(* IEC 61131-3 sources: daoli-st-library/DL_Base (part 10) *)

(* ---- FB_DL_CtudEx.st ---- *)
(*==============================================================================
 * 组件名称 (Component)  : FB_DL_CtudEx
 * 所属子库 (Sublibrary) : DL_Base
 * 当前版本 (Version)    : 1.0.0
 * 兼容性   (Platform)   : CODESYS 3.5 / TwinCAT 3 / 汇川 InoProShop / Machine Expert
 *                         仅依赖 Standard.library（R_TRIG），计数本体为库内显式
 *                         判界加减法（重实现最小化：一圈判界 + 加减 1）
 * 功能描述 (Function)   : 双向计数器（CTUD）防御包装。内部以两个 R_TRIG 标准实例
 *                         分别取 bCU / bCD 上升沿，CU/CD 同拍出现时按「净额抵消法」
 *                         取净值一次性施加（net = CU沿 − CD沿，同拍加减相消不误
 *                         动作）；优先级链 bRESET > bLOAD > 计数；PV 负值钳 0；
 *                         双向饱和不回绕（达 DINT 上/下限锁定并置故障码）。
 * 溯源     (Origin)     : IEC 61131-3 标准语义的道莅防御性实现
 *                         （接口语义由 IEC 61131-3 定义，clean-room 重写，
 *                         参考公开标准条款）
 * 码位     (Diag Codes) : 信息级 16#0001_0155（本件独占）：
 *                         nPV 为负值已钳 0 ／ CU/CD 同拍抵消（净变化 0）
 *                         故障级 16#0001_0226（本件独占）：
 *                         CV 达 DINT 上/下限饱和锁定（异常记录，绝不回绕）
 * 类型裁定 (Type Note)  : 码位段 16#0001_xxxx 为全库共享 32 位段，WORD 容量不足，
 *                         故 uDiag 采用 UDINT 承载（与库内 uErrorId : UDINT 惯例一致）
 * 边界声明 (Boundary)   : 本件是对标准 CTUD 的逐引脚等义防御包装（无双预设、无倒置
 *                         冻结扩展）；CTUD 全语义超集见 FB_DL_BidirectionalCounter，
 *                         两者在 MANUAL 中互引声明边界，不互相替代。
 * 依赖     (Depends)    : 无 DL_ 内部依赖；Standard.library: R_TRIG
 * 红线自检 (Redline)    : R1 ✓ 零全局变量与外部变量引用 ｜ R2 ✓ 零物理 IO 地址直写
 *                         R3 ✓ 纯 IEC 61131-3 ｜ R4 ✓ PV 钳位+DINT 双向判界防回绕
 *                         R5 ✓ 全变量中英双语同行注释 ｜ R6 N/A（无顺序状态机，见下）
 *                         R7 ✓ R_TRIG 实例主体无条件周期刷新
 * 说明     (Note)       : R6 标注 N/A —— 本组件为「复位/装载/计数」优先级时序
 *                         逻辑，非顺序步进状态机，无 CASE 可写；三态互斥由优先级
 *                         链（复位 > 装载 > 计数）显式保证，以本节说明替代
 *                         ELSE 兜底，符合"无状态机则标注 N/A"口径。
 * 防御行为声明 (Defense): ① CU/CD 同拍出现按「净额抵消法」处理：两沿同拍时
 *                           net = +1 − 1 = 0，本拍不动作并置信息码 16#0001_0155
 *                           （先加后减的顺序歧义被一次性净值施加天然规避）；
 *                         ② 优先级链写死：bRESET（电平）> bLOAD（电平）> 计数净值；
 *                           装载拍跳过计数（装载覆盖计数，与库内计数族口径一致）；
 *                         ③ nPV < 0 时钳位为 0 并置信息码 16#0001_0155
 *                           （负预置使 bQU 恒 TRUE，属组态错误提示）；
 *                         ④ 双向饱和不回绕：CV 达 DINT 上限 2147483647 停止递增、
 *                           达下限 −2147483648 停止递减，保持不变并置故障码
 *                           16#0001_0226（与标准 CTUD 的回绕行为差异点）；
 *                         ⑤ DINT 上/下限提为只读常量，禁魔法数。
 * 修订历史 (Revision)   :
 *   2026-11-16  v1.0.0  首版入库（R14 批 3 · T0 快车道）
 *============================================================================*)
FUNCTION_BLOCK FB_DL_CtudEx
VAR_INPUT
    bCU    : BOOL;  // 加计数脉冲输入（内部 R_TRIG 取沿） / Count-up pulse input (edge taken by internal R_TRIG)
    bCD    : BOOL;  // 减计数脉冲输入（内部 R_TRIG 取沿） / Count-down pulse input (edge taken by internal R_TRIG)
    bRESET : BOOL;  // 复位输入（电平，优先级最高），CV 清零 / Reset input (level, highest priority), clears CV
    bLOAD  : BOOL;  // 装载输入（电平，次高优先级），CV 装入钳位后 PV / Load input (level, second priority), loads clamped PV into CV
    nPV    : INT;   // 预置值 [个]，负值将被钳位为 0 / Preset value [count], negative values are clamped to 0
END_VAR
VAR_OUTPUT
    nCV   : DINT;   // 当前计数值 [个]，双向饱和不回绕 / Current count [count], saturates both ways without wrap
    bQU   : BOOL;   // 上计数到达输出，nCV >= 钳位后 nPV 时 TRUE / Upper done output, TRUE when nCV >= clamped nPV
    bQD   : BOOL;   // 下计数到达输出，nCV <= 0 时 TRUE / Lower done output, TRUE when nCV <= 0
    uDiag : UDINT;  // 诊断字，16#0001_0155=PV负钳0或同拍抵消，16#0001_0226=CV饱和，0=无事件 / Diag word, 16#0001_0155=PV clamped or same-scan cancel, 16#0001_0226=CV saturated, 0=no event
END_VAR
VAR
    fbCuTrig  : R_TRIG;  // 内建上升沿实例，取 bCU 计数脉冲 / Built-in R_TRIG instance for the count-up pulse
    fbCdTrig  : R_TRIG;  // 内建上升沿实例，取 bCD 计数脉冲 / Built-in R_TRIG instance for the count-down pulse
    nPVClamp  : DINT;    // 钳位后的预置值 [个]，用于装载与比较输出 / Clamped preset [count], used for load and compare outputs
    nNet      : INT;     // 本拍净计数额 [个]，加 1 / 减 1 / 0 抵消 / Net count delta this scan [count], plus one, minus one or zero
    xInit     : BOOL;    // 首扫初始化标志，FALSE=尚未完成上电初始化 / First-scan init flag, FALSE = power-on init not yet done
    nDintMax  : DINT := 2147483647;   // DINT 上限常量（只读语义，主体禁写）/ DINT upper-limit constant (read-only semantics, never written in body)
    nDintMin  : DINT := -2147483648;  // DINT 下限常量（只读语义，主体禁写）/ DINT lower-limit constant (read-only semantics, never written in body)
END_VAR

(*------------------------------------------------------------------------------
 * 段 1｜首扫初始化（历史教训④口径）：置于逻辑最前，首扫 CV=0、比较输出 FALSE
 *      First-scan init (lesson 4): placed at the very front, CV=0 and compare outputs FALSE on first scan
 *-----------------------------------------------------------------------------*)
IF NOT xInit THEN
    xInit    := TRUE;             // 置初始化完成标志 / Mark init as done
    nCV      := 0;                // 首扫计数值清零 [个] / Zero count on first scan [count]
    nPVClamp := 0;                // 首扫钳位预置清零 [个] / Zero clamped preset on first scan [count]
    nNet     := 0;                // 首扫净额清零 [个] / Zero net delta on first scan [count]
    uDiag    := 16#0000_0000;     // 首扫诊断字清零 / Clear diag word on first scan
END_IF

(*------------------------------------------------------------------------------
 * 段 2｜PV 域校验与钳位：nPV 负值钳 0 并置信息码 16#0001_0155
 *      PV domain check and clamp: negative nPV clamped to 0 with code 16#0001_0155
 *-----------------------------------------------------------------------------*)
IF nPV < 0 THEN
    nPVClamp := 0;                // 负预置钳位为 0 [个] / Clamp negative preset to 0 [count]
    uDiag    := 16#0001_0155;     // 信息码：nPV 负值已钳 0 / Informational: negative nPV clamped to 0
ELSE
    nPVClamp := nPV;              // 域内直通 [个] / In-domain pass-through [count]
    uDiag    := 16#0000_0000;     // 无诊断事件，清码 / No diag event, clear code
END_IF

(*------------------------------------------------------------------------------
 * 段 3｜无条件刷新区（红线 R7）：两个 R_TRIG 实例严禁进入任何 IF / CASE 分支
 *      Unconditional refresh zone (red line R7): no instance call inside IF / CASE
 *-----------------------------------------------------------------------------*)
fbCuTrig(CLK := bCU);  // 每扫描周期无条件取 bCU 上升沿 / Take bCU rising edge unconditionally every scan
fbCdTrig(CLK := bCD);  // 每扫描周期无条件取 bCD 上升沿 / Take bCD rising edge unconditionally every scan

(*------------------------------------------------------------------------------
 * 段 4｜净额抵消仲裁（防御声明①）：CU/CD 同拍时 net = 0，同拍加减相消不误动作；
 *      净额一次性施加，杜绝「先加后减还是先减后加」的平台顺序歧义
 *      Net-amount arbitration (defense note 1): same-scan CU and CD edges cancel
 *      to net zero; the net value is applied once, eliminating order ambiguity
 *-----------------------------------------------------------------------------*)
IF fbCuTrig.Q AND fbCdTrig.Q THEN
    nNet  := 0;                   // 同拍双向抵消，净变化 0 [个] / Same-scan bidirectional cancel, net zero [count]
    uDiag := 16#0001_0155;        // 信息码：同拍抵消已记录 / Informational: same-scan cancel recorded
ELSIF fbCuTrig.Q THEN
    nNet := 1;                    // 仅加沿，净额 +1 [个] / Up edge only, net plus one [count]
ELSIF fbCdTrig.Q THEN
    nNet := -1;                   // 仅减沿，净额 -1 [个] / Down edge only, net minus one [count]
ELSE
    nNet := 0;                    // 无计数沿，净额 0 [个] / No count edge, net zero [count]
END_IF

(*------------------------------------------------------------------------------
 * 段 5｜计数主体（优先级链 bRESET > bLOAD > 计数，防御声明②）：
 *      双向饱和判界先行——达 DINT 上/下限锁定并置故障码，绝不回绕
 *      Count body (priority chain bRESET > bLOAD > count, defense note 2):
 *      both-direction saturation checked before the update, no wrap ever
 *-----------------------------------------------------------------------------*)
IF bRESET THEN
    nCV := 0;                     // 复位清零计数值 [个] / Reset clears count [count]
ELSIF bLOAD THEN
    nCV := nPVClamp;              // 装载钳位后预置 [个]，本拍跳过计数 / Load clamped preset [count], counting skipped this scan
ELSIF nNet = 1 THEN
    IF nCV < nDintMax THEN
        nCV := nCV + 1;           // 域内递增 1 [个] / In-domain increment by 1 [count]
    ELSE
        uDiag := 16#0001_0226;    // 故障码：CV 上限饱和锁定，不回绕 / Fault: CV upper-limit saturation, no wrap
    END_IF
ELSIF nNet = -1 THEN
    IF nCV > nDintMin THEN
        nCV := nCV - 1;           // 域内递减 1 [个] / In-domain decrement by 1 [count]
    ELSE
        uDiag := 16#0001_0226;    // 故障码：CV 下限饱和锁定，不回绕 / Fault: CV lower-limit saturation, no wrap
    END_IF
END_IF

(*------------------------------------------------------------------------------
 * 段 6｜比较输出：按 IEC CTUD 语义 QU = CV >= PV、QD = CV <= 0
 *      （PV 钳 0 时 bQU 恒 TRUE，属组态提示范畴，见头注释防御声明③）
 *      Compare outputs: per IEC CTUD semantics QU = CV >= PV and QD = CV <= 0
 *      (bQU always TRUE when PV clamped to 0, a configuration hint, defense note 3)
 *-----------------------------------------------------------------------------*)
bQU := (nCV >= nPVClamp);  // 上计数到达比较 [个] / Upper done comparison [count]
bQD := (nCV <= 0);         // 下计数到达比较 [个] / Lower done comparison [count]
END_FUNCTION_BLOCK

(* ---- FB_DL_CtuEx.st ---- *)
(*==============================================================================
 * 组件名称 (Component)  : FB_DL_CtuEx
 * 所属子库 (Sublibrary) : DL_Base
 * 当前版本 (Version)    : 1.0.0
 * 兼容性   (Platform)   : CODESYS 3.5 / TwinCAT 3 / 汇川 InoProShop / Machine Expert
 *                         仅依赖 Standard.library（R_TRIG），计数本体为库内显式
 *                         判界加减法（重实现最小化：仅一圈判界 + 加 1）
 * 功能描述 (Function)   : 加计数器防御包装。内部以 R_TRIG 标准实例产计数脉冲，
 *                         计数本体采用显式判界加法实现 CV 饱和不回绕（达 DINT
 *                         上限锁定并置诊断码）；复位优先级 bRESET > bCU。
 * 溯源     (Origin)     : IEC 61131-3 标准语义的道莅防御性实现
 *                         （接口语义由 IEC 61131-3 定义，clean-room 重写，
 *                         参考公开标准条款）
 * 码位     (Diag Codes) : 信息级占用区间 16#0001_0153（本件独占，仅此一码，
 *                         双事件共用一类码）
 *                         16#0001_0153 = nPV 为负值已钳 0 ／ CV 达 DINT 上限
 *                         饱和锁定（信息级，饱和是正常防御行为，不置故障）
 * 类型裁定 (Type Note)  : 码位段 16#0001_xxxx 为全库共享 32 位段，WORD 容量不足，
 *                         故 uDiag 采用 UDINT 承载（与库内 uErrorId : UDINT 惯例一致）
 * 依赖     (Depends)    : 无 DL_ 内部依赖；Standard.library: R_TRIG
 * 红线自检 (Redline)    : R1 ✓ 零全局变量与外部变量引用 ｜ R2 ✓ 零物理 IO 地址直写
 *                         R3 ✓ 纯 IEC 61131-3 ｜ R4 ✓ PV 钳位+DINT 上限判界防回绕
 *                         R5 ✓ 全变量中英双语同行注释 ｜ R6 N/A（无顺序状态机，见下）
 *                         R7 ✓ R_TRIG 实例主体无条件周期刷新
 * 说明     (Note)       : R6 标注 N/A —— 本组件为「复位/计数」双态时序逻辑，
 *                         非顺序步进状态机，无 CASE 可写；两态互斥由优先级链
 *                         （复位 > 计数）显式保证，以本节说明替代 ELSE 兜底，
 *                         符合"无状态机则标注 N/A"口径。
 * 防御行为声明 (Defense): ① nPV < 0 时钳位为 0 并置信息码 16#0001_0153
 *                           （负预置在本包装下使 bQ 恒 TRUE，属组态错误提示）；
 *                         ② 上溢饱和不回绕：CV 达 DINT 上限 2147483647 后停止
 *                           递增、保持不变并置信息码（与标准 CTU 的 DINT 回绕
 *                           行为差异点，饱和是正常防御行为）；
 *                         ③ 优先级链写死：bRESET（电平）> bCU 计数脉冲；
 *                         ④ 内部状态量写入点排序审计（历史教训⑦）：PV 钳位段
 *                           与计数段对 uDiag 只写同一码值 16#0001_0153，不存在
 *                           复位类与置位类竞态，排序安全；
 *                         ⑤ DINT 上限提为只读常量 nDintMax，禁魔法数。
 * 修订历史 (Revision)   :
 *   2026-11-16  v1.0.0  首版入库（R14 批 2 · T0 快车道）
 *============================================================================*)
FUNCTION_BLOCK FB_DL_CtuEx
VAR_INPUT
    bCU    : BOOL;  // 加计数脉冲输入（内部 R_TRIG 取沿） / Count-up pulse input (edge taken by internal R_TRIG)
    bRESET : BOOL;  // 复位输入（电平，优先级最高），CV 清零 / Reset input (level, highest priority), clears CV
    nPV    : INT;   // 预置值 [个]，负值将被钳位为 0 / Preset value [count], negative values are clamped to 0
END_VAR
VAR_OUTPUT
    nCV   : DINT;   // 当前计数值 [个]，达上限饱和不回绕 / Current count [count], saturates at upper limit without wrap
    bQ    : BOOL;   // 计数到达输出，nCV >= 钳位后 nPV 时 TRUE / Done output, TRUE when nCV >= clamped nPV
    uDiag : UDINT;  // 诊断字，16#0001_0153=nPV 负钳 0 或 CV 上限饱和，0=无事件 / Diag word, 16#0001_0153=negative nPV clamped or CV upper saturation, 0=no event
END_VAR
VAR
    fbCuTrig  : R_TRIG;  // 内建上升沿实例，产计数脉冲 / Built-in R_TRIG instance, generates the count pulse
    nPVClamp  : DINT;    // 钳位后的预置值 [个]，用于比较输出 / Clamped preset [count], used for the compare output
    nDintMax  : DINT := 2147483647;  // DINT 上限常量（只读语义，主体禁写）/ DINT upper-limit constant (read-only semantics, never written in body)
    xInit     : BOOL;    // 首扫初始化标志，FALSE=尚未完成上电初始化 / First-scan init flag, FALSE = power-on init not yet done
END_VAR

(*------------------------------------------------------------------------------
 * 段 1｜首扫初始化（历史教训④口径）：置于逻辑最前，首扫 CV=0、bQ=FALSE
 *      First-scan init (lesson 4): placed at the very front, CV=0 and bQ=FALSE on first scan
 *-----------------------------------------------------------------------------*)
IF NOT xInit THEN
    xInit    := TRUE;    // 置初始化完成标志 / Mark init as done
    nCV      := 0;       // 首扫计数值清零 [个] / Zero count on first scan [count]
    nPVClamp := 0;       // 首扫钳位预置清零 [个] / Zero clamped preset on first scan [count]
    uDiag    := 16#0000_0000;  // 首扫诊断字清零 / Clear diag word on first scan
END_IF

(*------------------------------------------------------------------------------
 * 段 2｜PV 域校验与钳位（历史教训⑨）：nPV 负值钳 0 并置信息码
 *      PV domain check and clamp (lesson 9): negative nPV clamped to 0 with code
 *-----------------------------------------------------------------------------*)
IF nPV < 0 THEN
    nPVClamp := 0;            // 负预置钳位为 0 [个] / Clamp negative preset to 0 [count]
    uDiag    := 16#0001_0153;  // 信息码：nPV 负值已钳 0 / Informational: negative nPV clamped to 0
ELSE
    nPVClamp := nPV;          // 域内直通 [个] / In-domain pass-through [count]
    uDiag    := 16#0000_0000;  // 无诊断事件，清码 / No diag event, clear code
END_IF

(*------------------------------------------------------------------------------
 * 段 3｜无条件刷新区（红线 R7）：R_TRIG 实例严禁进入任何 IF / CASE 分支
 *      Unconditional refresh zone (red line R7): no instance call inside IF / CASE
 *-----------------------------------------------------------------------------*)
fbCuTrig(CLK := bCU);  // 每扫描周期无条件取 bCU 上升沿 / Take bCU rising edge unconditionally every scan

(*------------------------------------------------------------------------------
 * 段 4｜计数主体（优先级链 bRESET > bCU）：复位电平优先，计数沿次之；
 *      上溢判界先行——CV 达 DINT 上限停止递增并置饱和码，绝不回绕
 *      Count body (priority chain bRESET > bCU): reset level first, count edge
 *      second; overflow boundary checked before increment, no wrap ever
 *-----------------------------------------------------------------------------*)
IF bRESET THEN
    nCV := 0;   // 复位清零计数值 [个] / Reset clears count [count]
ELSIF fbCuTrig.Q THEN
    IF nCV < nDintMax THEN
        nCV := nCV + 1;           // 域内递增 1 [个] / In-domain increment by 1 [count]
    ELSE
        uDiag := 16#0001_0153;    // 信息码：CV 上限饱和锁定，不回绕 / Informational: CV upper-limit saturation, no wrap
    END_IF
END_IF

(*------------------------------------------------------------------------------
 * 段 5｜比较输出：按 IEC CTU 语义 Q = CV >= PV（PV 钳 0 时恒 TRUE，属组态
 *      提示范畴，见头注释防御声明①）
 *      Compare output: per IEC CTU semantics Q = CV >= PV (always TRUE when
 *      PV clamped to 0, a configuration hint, see defense note 1)
 *-----------------------------------------------------------------------------*)
bQ := (nCV >= nPVClamp);  // 计数到达比较 [个] / Done comparison [count]
END_FUNCTION_BLOCK

(* ---- FB_DL_CycleBarrierGate.st ---- *)
(*==============================================================================
 * 组件名称 (Component)  : FB_DL_CycleBarrierGate
 * 所属子库 (Sublibrary) : DL_Base
 * 当前版本 (Version)    : 1.0.0
 * 兼容性 (Platform)     : CODESYS 3.5+ / TwinCAT 3 / 汇川 InoProShop / 施耐德 Machine Expert
 *                         仅依赖 Standard.library（TON），零厂商私有库
 * 功能描述 (Function)   : 多设备同周期相位会合闸（集合点原语）。nMemberCount 个
 *                         成员各自上报就绪电平（abMemberReady），全部就绪时
 *                         bGateOpen 单拍放行并清到达掩码；若在 tWindow 内未能
 *                         全员到齐 → bBarrierTimeout 置位并锁存滞留成员掩码
 *                         （诊断用），需 bAck 确认后重新等待。产线多工站同拍
 *                         会合、多轴同步起点、批处理工序齐套场景。
 * 来源标签 (Origin)     : 自研线（IEC 61131-3 标准语义的道莅防御性实现，clean-room）
 * 分工声明 (Pairing)    : CycleBarrierGate（会合闸，本件）↔ FB_DL_SemaMutex（互斥，
 *                         既有件）：本件管「全员齐套统一放行」（AND 集合点），
 *                         不管「资源独占互斥」；SemaMutex 管令牌互斥，不做
 *                         齐套判据（R298 属主边界）。
 * 输出语义 (Fallback)   : 【R191】bEnable = FALSE → bGateOpen 强制 FALSE（放行
 *                         是安全相关动作，失能必须收敛），到达掩码冻结保持；
 *                         eFault 相 → bGateOpen 保持 FALSE，bError = TRUE。
 * 组态闸 (Config gate)  : nMemberCount < 2 或 > 16（集合点无意义/超容量）或
 *                         tWindow <= T#0S → 故障锁存。
 * 码位     (Codes)      : 按 R297 范式零 16# 码位硬编码；错误出口 BOOL+ENUM(eCause)，
 *                         码位待主控收口统一派号。
 * 红线自检 (Redline)    : 7 项红线已自检：R1 零全局 ✓｜R2 零物理地址 ✓｜R3 纯 IEC ✓
 *                         R4 组态闸/数组下标钳位 ✓｜R5 双语同行注释 ✓
 *                         R6 CASE 带 ELSE 兜底迁 eFault ✓｜R7 TON 段 0 无条件刷新 ✓
 * 验收向量 (Acceptance) : V1 4 成员全员就绪 → bGateOpen 单拍 TRUE 且掩码清零；
 *                         V2 窗口到时仅 3/4 就绪 → bBarrierTimeout=TRUE，
 *                         uLatchedMask 指示滞留成员位；
 *                         V3 nMemberCount=1 → eFault 锁存。
 * 修订历史 (Revision)   : 2026-11-20  v1.0.0  R49 首版（批 2 · 序号 6）
 *==============================================================================*)
TYPE E_DL_CbgState :
(
    eIdle    := 0,                           (* 待启动（闸门关闭） / Idle, gate closed *)
    eWait    := 10,                          (* 等待全员就绪 / Waiting for all members *)
    eTimeout := 20,                          (* 窗口超时滞留，等确认 / Timeout stranded, awaiting ack *)
    eFault   := 90                           (* 故障锁存相 / Fault latched phase *)
);
END_TYPE

TYPE E_DL_CbgCause :
(
    eNone       := 0,                        (* 无故障成因 / No cause *)
    eCfgIllegal := 1,                        (* 组态非法：成员数/窗口越域 / Illegal config *)
    ePhaseBad   := 2                         (* 非法相位兜底 / Illegal phase fallback *)
);
END_TYPE

FUNCTION_BLOCK FB_DL_CycleBarrierGate
VAR_INPUT
    abMemberReady : ARRAY[1..16] OF BOOL;    (* 成员就绪电平数组（按位消费前 nCount 个）[-] / Member ready levels *)
    nMemberCount  : INT := 4;                (* 参与会合成员数，域 2..16 [个] / Member count, domain 2..16 *)
    tWindow       : TIME := T#5S;            (* 全员到齐窗口保持时长 [ms] / All-arrive window hold time *)
    bStart        : BOOL := FALSE;           (* 会合启动电平，TRUE 开始等待 / Barrier start level *)
    bAck          : BOOL := FALSE;           (* 超时确认，上升沿清滞留掩码并重新等待 [-] / Timeout ack, rising edge clears strand mask *)
    bEnable       : BOOL := TRUE;            (* 会合闸使能，FALSE 时放行强制收敛 [-] / Gate enable *)
    bReset        : BOOL := FALSE;           (* 复位命令，上升沿清全部内部状态 [-] / Reset command *)
END_VAR
VAR_OUTPUT
    bGateOpen        : BOOL;                 (* 放行单拍位（全员到齐拍置位）[-] / Gate-open single-scan pulse *)
    uArrivedMask     : UDINT;                (* 当前已到达成员位掩码（实时）[-] / Current arrived member bitmask *)
    uLatchedMask     : UDINT;                (* 超时滞留成员位掩码（锁存至 bAck）[-] / Stranded member bitmask latched until ack *)
    nArrivedCnt      : INT;                  (* 已到达成员数（实时）[个] / Arrived member count *)
    bBarrierTimeout  : BOOL;                 (* 窗口超时锁存位（bAck 清）[-] / Window timeout latch, cleared by ack *)
    eState           : E_DL_CbgState;        (* 状态出口 / State outlet *)
    eCause           : E_DL_CbgCause;        (* 故障成因出口（R190 归因唯一） / Fault cause outlet *)
    bError           : BOOL;                 (* 故障锁存标志 [-] / Fault latch flag *)
END_VAR
VAR
    _eState   : E_DL_CbgState := E_DL_CbgState.eIdle;     (* 内部相位（CASE 唯一写入目标） / Internal phase *)
    _eCause   : E_DL_CbgCause := E_DL_CbgCause.eNone;     (* 故障成因锁存量 / Latched cause *)
    rtAck     : R_TRIG;                     (* 确认沿实例，段 0 无条件调用 / Ack edge instance *)
    rtReset   : R_TRIG;                     (* 复位沿实例，段 0 无条件调用 / Reset edge instance *)
    tonWindow : TON;                        (* 到齐窗口计时，IN 由相位派生 / Window timer *)
    _nArrived : INT;                        (* 到达计数当拍派生量 [个] / Arrived count derived this scan *)
    _uMask    : UDINT;                      (* 到达掩码当拍派生量 / Arrived bitmask derived *)
    _bAllArr  : BOOL;                       (* 全员到齐当拍判据 / All-arrived verdict *)
    _i        : INT;                        (* 成员扫描游标（每趟重置，R227）[-] / Member scan cursor *)
    _bFault   : BOOL;                       (* 故障锁存位 / Latched fault bit *)
    _bCfgBad  : BOOL;                       (* 组态非法当拍量 / Illegal config this scan *)
END_VAR

(* —— 段 0：当拍判据派生 + 实例无条件刷新（R228A） —— *)
_bCfgBad := (nMemberCount < 2) OR (nMemberCount > 16) OR (tWindow <= T#0S);   (* 组态闸 / Config gate *)
rtAck(CLK := bAck);                                                          (* 确认沿每拍必调 / Ack edge every scan *)
rtReset(CLK := bReset);                                                      (* 复位沿每拍必调 / Reset edge every scan *)
tonWindow(IN := _eState = E_DL_CbgState.eWait, PT := tWindow);               (* 窗口计时随相位派生 / Window timer phase-derived *)
_uMask := 0;                                                                 (* 掩码派生量清零重扫 / Mask derived recompute *)
_nArrived := 0;                                                              (* 到达计数清零重扫 / Count derived recompute *)
_i := 1;                                                                     (* 游标起头显式重置（R227） / Cursor reset *)
WHILE _i <= nMemberCount DO                                                  (* 只扫前 nCount 个成员（容量内，无越界） / Scan first nCount members *)
    _uMask := _uMask + _uMask;                                               (* 先整体左移一位（UDINT 域 16 成员最大 2^16 无溢出，免 SHL 移位量归一，R295） / Shift left first *)
    IF abMemberReady[_i] THEN
        _uMask := _uMask + 1;                                                (* 后置位最低位：成员 i 落于位 i-1（自证向量：i=1→bit0，i=2→bit1） / Then set LSB: member i maps to bit i-1 *)
        _nArrived := _nArrived + 1;                                          (* 到达计数 / Arrived count *)
    END_IF
    _i := _i + 1;                                                            (* 游标递进 / Cursor advance *)
END_WHILE
_bAllArr := (_nArrived >= nMemberCount);                                     (* 全员到齐判据（整数等值域合法） / All-arrived verdict *)

(* —— 段 1：单拍量预清零（R107） —— *)
bGateOpen := FALSE;                                                          (* 放行单拍位预清，唯一分支置位 / Gate pulse preset *)

(* —— 段 2：复位沿处理（作用域：清故障 + 清掩码锁存 + 清超时 + 迁 eIdle，R283 逐项声明） —— *)
IF rtReset.Q THEN
    _bFault := FALSE;                                                       (* 清故障锁存 / Clear fault *)
    _eCause := E_DL_CbgCause.eNone;                                         (* 清成因 / Clear cause *)
    uLatchedMask := 0;                                                      (* 清滞留掩码锁存 / Clear strand mask *)
    bBarrierTimeout := FALSE;                                               (* 清超时锁存 / Clear timeout latch *)
    _eState := E_DL_CbgState.eIdle;                                         (* 迁待启动相 / Back to idle *)
END_IF

(* —— 段 3：组态闸故障锁存（R45 配对；锁存至复位沿，R189） —— *)
IF _bCfgBad AND NOT _bFault THEN
    _bFault := TRUE;                                                        (* 锁存故障位 / Latch fault *)
    _eCause := E_DL_CbgCause.eCfgIllegal;                                   (* 成因：组态非法 / Cause: illegal config *)
    _eState := E_DL_CbgState.eFault;                                        (* 同步迁故障相 / Migrate to fault *)
END_IF

(* —— 段 4：CASE 主状态机（ELSE 兜底迁 eFault，红线 6） —— *)
CASE _eState OF
    E_DL_CbgState.eIdle:                                                    (* 待启动相 / Idle *)
        IF bStart AND bEnable AND NOT _bFault THEN
            _eState := E_DL_CbgState.eWait;                                 (* 启动进入等待 / Start enters wait *)
        END_IF
    E_DL_CbgState.eWait:                                                    (* 等待全员相 / Wait *)
        IF NOT bEnable OR NOT bStart THEN                                   (* 启动撤销回待机 / Start withdrawn *)
            _eState := E_DL_CbgState.eIdle;                                 (* 回待启动 / Back to idle *)
        ELSIF _bAllArr THEN                                                 (* 全员到齐 / All arrived *)
            bGateOpen := TRUE;                                              (* 放行单拍脉冲 / Gate pulse *)
            _eState := E_DL_CbgState.eIdle;                                 (* 本周期会合完成回待机（每周期重新集合语义） / Round complete, re-convene next cycle *)
        ELSIF tonWindow.Q THEN                                              (* 窗口到时未齐 / Window expired *)
            uLatchedMask := _uMask;                                         (* 锁存滞留掩码（诊断：值为 1 的位 = 已到，0 的位 = 滞留） / Latch strand mask *)
            bBarrierTimeout := TRUE;                                        (* 超时锁存至 bAck / Timeout latch *)
            _eState := E_DL_CbgState.eTimeout;                              (* 迁超时相 / Enter timeout *)
        END_IF
    E_DL_CbgState.eTimeout:                                                 (* 超时滞留相 / Timeout *)
        IF rtAck.Q THEN                                                     (* 确认沿：清锁存重新等待 / Ack: clear latch, re-wait *)
            uLatchedMask := 0;                                              (* 清滞留掩码 / Clear strand mask *)
            bBarrierTimeout := FALSE;                                       (* 清超时锁存 / Clear timeout latch *)
            _eState := E_DL_CbgState.eWait;                                 (* 重新等待（eWait 相退出条件：事件沿 + 状态清除双条件） / Re-enter wait *)
        ELSIF NOT bEnable OR NOT bStart THEN
            _eState := E_DL_CbgState.eIdle;                                 (* 启动撤销亦可退出（第二退出条件） / Start withdrawn exit *)
        END_IF
    E_DL_CbgState.eFault:                                                   (* 故障相：仅复位沿出 / Fault *)
        ;                                                                   (* 锁存回放（R28） / Replay from latch *)
    ELSE                                                                    (* 非法相位兜底迁安全态 / Illegal phase fallback *)
        _eState := E_DL_CbgState.eFault;                                    (* 迁故障相 / To fault *)
        _bFault := TRUE;                                                    (* 同步锁存 / Latch *)
        _eCause := E_DL_CbgCause.ePhaseBad;                                 (* 成因：非法相位 / Cause: illegal phase *)
END_CASE

(* —— 段 5：出口映射（bError/eState 同源，R191） —— *)
uArrivedMask := _uMask;                                                     (* 到达掩码实时镜像 / Arrived mask mirror *)
nArrivedCnt := _nArrived;                                                   (* 到达计数实时镜像 / Arrived count mirror *)
bError := _bFault;                                                          (* 故障标志镜像 / Fault flag mirror *)
eState := _eState;                                                          (* 状态出口 / State outlet *)
eCause := _eCause;                                                          (* 成因出口 / Cause outlet *)
END_FUNCTION_BLOCK

(* ---- FB_DL_CycleTimeMeasure.st ---- *)
(*==============================================================================
 * 组件名称 (Component)  : FB_DL_CycleTimeMeasure
 * 所属子库 (Sublibrary) : DL_Base
 * 当前版本 (Version)    : 1.0.0
 * 兼容性   (Platform)   : CODESYS 3.5 / TwinCAT 3 / 汇川 InoProShop / Machine Expert
 *                         仅依赖 Standard.library（R_TRIG），零平台时刻函数
 * 功能描述 (Function)   : 任务扫描周期统计（最近 / 最小 / 最大 / 平均 / 样本数）。
 *                         本块自身不读取任何平台时刻，时间增量由调用方以输入引脚注入，
 *                         因此零平台依赖、三平台可编译，平台差异被关在调用方一处。
 *                         零增量与超上限增量一律拒收并告警，避免垃圾样本污染极值；
 *                         窗内首个有效样本同时初始化最小值与最大值（不得以 0 当初始值）；
 *                         样本数达上限自动重开统计窗并告警（无符号累计上限保护）。
 * 开源溯源 (Origin)     : 原创实现。指标口径（最近/最小/最大/平均/样本数）参照
 *                         工业界周期监控块的通用输出集合；时间注入设计为本库对
 *                         平台时刻函数依赖的主动拒绝方案，未复制任何源码。
 * 本文件内含       : FB    FB_DL_CycleTimeMeasure（单 POU，无配套类型）
 * 依赖     (Depends)    : 无 DL_ 内部依赖；Standard.library: R_TRIG
 * 红线自检 (Redline)    : R1 ✓ 禁用全局存储与物理寻址 ｜ R2 ✓ 无地址直写
 *                         R3 ✓ 纯 IEC 61131-3，零平台时刻函数 ｜ R4 ✓ 除零双保险 + 数据拒收 + 窗滚动
 *                         R5 ✓ 全变量中英双语同行注释 ｜ R6 N/A（纯统计累加，无跨周期状态转移）
 *                         R7 ✓ R_TRIG 主体最前部无条件刷新 ｜ R8 ✓ 上限与阈值全常量化
 *
 * 【调用方契约 / Caller contract（边界 B8）】
 *   调用方须在同一任务内以"当前系统时刻 − 上周期系统时刻"得到毫秒增量后注入本引脚；
 *   首扫须跳过或注入一个已知有效值，否则 0 增量会被本块按无效数据处理并告警。
 *   本块不做任何时刻获取、不做跨任务共享，一个任务一个实例。
 *
 * 修订历史 (Revision)   :
 *   2026-11-14  v1.0.0  首版入库（Phase 1 第二轮 · Level 0 批次 A）
 *============================================================================*)
FUNCTION_BLOCK FB_DL_CycleTimeMeasure
VAR_INPUT
    uDeltaTimeMs : UDINT;              // 本任务周期实际耗时 [ms]，调用方注入 / Actual cycle time in ms, caller-provided
    bCapture     : BOOL := TRUE;       // TRUE = 本周期计入统计 / TRUE = include this cycle in statistics
    bReset       : BOOL;               // 上升沿清空全部统计 / Rising edge clears statistics
END_VAR
VAR_OUTPUT
    uCycleLast   : UDINT;              // 最近一个有效周期 [ms] / Last valid cycle time [ms]
    uCycleMin    : UDINT;              // 统计窗内最小周期 [ms] / Minimum in window [ms]
    uCycleMax    : UDINT;              // 统计窗内最大周期 [ms] / Maximum in window [ms]
    fCycleMean   : REAL;               // 统计窗内平均周期 [ms] / Mean in window [ms]
    nSampleCount : UDINT;              // 统计窗内样本数 [个] / Sample count in window [count]
    uErrorId     : UDINT;              // 故障码，0 = 无故障 / Error code, 0 = no error
END_VAR
VAR
    uSumMs       : UDINT;              // 窗内累计耗时总和 [ms] / Accumulated sum in window [ms]
    fbTrigReset  : R_TRIG;             // 复位上升沿检测实例 / Reset rising edge detector instance
    bDeltaValid  : BOOL;               // 本周期增量有效性判定结果 / Current-cycle delta validity result
END_VAR
VAR CONSTANT
    DL_CYC_SAMPLE_MAX : UDINT := 1000000;   // 统计窗样本上限，达限自动重开窗 / Window sample cap, auto reopen at limit
    DL_CYC_DELTA_MAX  : UDINT := 3600000;   // 单周期合理上限 [ms]，超限视为无效数据 / Sanity cap per cycle [ms]
END_VAR

(*------------------------------------------------------------------------------
 * 段 1｜无条件刷新区（红线 R7）：复位沿实例位于主体最前部，严禁进入 IF / CASE
 *      Unconditional refresh zone: the reset edge instance runs at the very top
 *-----------------------------------------------------------------------------*)
fbTrigReset(CLK := bReset);

(*------------------------------------------------------------------------------
 * 段 2｜故障码本周期清零：错误码是"当前周期事实"，不是跨周期锁存量
 *      Error code is cleared every scan: it reports the current cycle only
 *-----------------------------------------------------------------------------*)
uErrorId := 16#0000_0000;

(*------------------------------------------------------------------------------
 * 段 3｜复位语义（边界 B7）：全部统计量归零，下一有效样本重新初始化极值
 *      Reset: clear every statistic, the next valid sample re-initialises extremes
 *-----------------------------------------------------------------------------*)
IF fbTrigReset.Q THEN
    uCycleLast   := UDINT#0;
    uCycleMin    := UDINT#0;
    uCycleMax    := UDINT#0;
    fCycleMean   := 0.0;
    nSampleCount := UDINT#0;
    uSumMs       := UDINT#0;
END_IF

(*------------------------------------------------------------------------------
 * 段 4｜增量合法性判定（边界 B2/B3）：0 表示调用方没取到时间，不是 0ms 快周期
 *      Delta validity: zero means the caller failed to read time, not a 0 ms cycle
 *      超上限增量同样拒收，防止取错基准产生的垃圾样本把 min / max 永久污染
 *      Over-limit deltas are rejected too, so a wrong time base cannot poison extremes
 *-----------------------------------------------------------------------------*)
IF (uDeltaTimeMs = UDINT#0) OR (uDeltaTimeMs > DL_CYC_DELTA_MAX) THEN
    bDeltaValid := FALSE;
    uErrorId    := 16#0001_0008;
ELSE
    bDeltaValid := TRUE;
END_IF

(*------------------------------------------------------------------------------
 * 段 5｜统计窗滚动（边界 B6）：样本数达上限先重开窗再采集，避免无符号累计失控
 *      Window rolling: reopen the window before sampling when the cap is reached
 *      重开窗保留 uCycleLast（HMI 上最近值不能跳变），min / max / sum / count 清零
 *      uCycleLast is preserved across a reopen so the HMI last-value does not jump
 *-----------------------------------------------------------------------------*)
IF nSampleCount >= DL_CYC_SAMPLE_MAX THEN
    uCycleMin    := UDINT#0;
    uCycleMax    := UDINT#0;
    fCycleMean   := 0.0;
    nSampleCount := UDINT#0;
    uSumMs       := UDINT#0;
    uErrorId     := 16#0001_0007;
END_IF

(*------------------------------------------------------------------------------
 * 段 6｜采样与极值更新（边界 B4）：首样本同时写入最小与最大值
 *      Sampling and extremes: the first valid sample initialises both min and max
 *      以 0 当初始值会让最小值永远是 0——经典缺陷，此处以计数为零作首样本判据
 *      Initialising with zero would pin the minimum at zero forever
 *-----------------------------------------------------------------------------*)
IF bDeltaValid AND bCapture THEN

    uCycleLast := uDeltaTimeMs;

    IF nSampleCount = UDINT#0 THEN
        (* 首样本：双极值同时落位，不存在"初值 0"参与比较 *)
        (* First sample: both extremes take the value, no zero seed participates *)
        uCycleMin := uDeltaTimeMs;
        uCycleMax := uDeltaTimeMs;
    ELSE
        IF uDeltaTimeMs < uCycleMin THEN
            uCycleMin := uDeltaTimeMs;
        END_IF
        IF uDeltaTimeMs > uCycleMax THEN
            uCycleMax := uDeltaTimeMs;
        END_IF
    END_IF

    uSumMs       := uSumMs + uDeltaTimeMs;
    nSampleCount := nSampleCount + UDINT#1;

END_IF

(*------------------------------------------------------------------------------
 * 段 7｜平均值输出（边界 B5）：除零双保险——计数判零 + 除数显式转换
 *      Mean output: dual divide-by-zero protection before the conversion
 *-----------------------------------------------------------------------------*)
IF nSampleCount > UDINT#0 THEN
    fCycleMean := UDINT_TO_REAL(uSumMs) / UDINT_TO_REAL(nSampleCount);
ELSE
    fCycleMean := 0.0;
END_IF
END_FUNCTION_BLOCK

(* ---- FB_DL_DebounceBank.st ---- *)
(*==============================================================================
 * 组件名称 (Component)  : FB_DL_DebounceBank
 * 所属子库 (Sublibrary) : DL_Base
 * 当前版本 (Version)    : 1.0.0
 * 兼容性   (Platform)   : CODESYS 3.5+ / TwinCAT 3 / 汇川 InoProShop / 施耐德 Machine Expert
 *                         仅依赖 Standard.library（TON），零厂商私有库
 * 功能描述 (Function)   : 16 路独立去抖库：每通道双阈值去抖（上升沿经 tRise
 *                         确认置 TRUE、下降沿经 tFall 确认回 FALSE，确认窗内
 *                         输出保持原态），每通道独立 TON 对（tonRise/tonFall），
 *                         全部实例主体无条件周期刷新（R6，禁止 IF 内调用）。
 *                         通道数 nChanCnt 钳位 1~16，越界钳位并置信息码
 *                         eCfgClamp；有效通道数之外的通道输出恒 FALSE。
 * 接口     (Interface)  : 输入 abRaw 16 路原始输入、aRise 16 路上升确认时间、
 *                         aFall 16 路下降确认时间、nChanCnt 有效通道数（钳位
 *                         1~16）；输出 abDeb 16 路去抖输出、bStable 全通道
 *                         稳定指示（全部通道当前不在确认窗内）、eErrCode
 *                         信息码、bError 故障标志（本件钳位走信息级，
 *                         bError 恒 FALSE，契约位保留）。
 * 边界     (Boundary)   : ① **属主边界（写死）：本件只做逐通道去抖，不判信号
 *                         语义、不做脉冲整形**；最小脉宽滤除归
 *                         `FB_DL_MinPulseWidthFilter`。
 *                         ② 32 个 TON 实例按 0..15 定长数组声明，FOR 循环
 *                         无条件调用（界宽常量，无死循环、无越界路径）。
 *                         ③ 双阈值语义：abDeb[i]=TRUE 当且仅当 tonRise[i].Q；
 *                          =FALSE 当 tonFall[i].Q（IN := NOT abRaw[i]）；两窗
 *                         均未到时输出保持上拍（互斥保持，无抖动带）。
 *                         ④ nChanCnt < 1 或 > 16：钳位到 [1,16] 并置信息码
 *                         eCfgClamp（规格指定钳位语义，不锁存故障）；有效域外
 *                         通道（i >= nChanCnt）输出强制 FALSE 且不参与 bStable。
 *                         ⑤ 时间引脚 <= T#0S 的通道按 0 处理（去抖直通：
 *                         输出跟随原始信号，TON PT=0 当拍到）。
 *                         ⑥ 零全局耦合（无 GVL / VAR_EXTERNAL / 物理地址）。
 * 分工声明 (Scope)      : 与 `FB_DL_SignalDebounce`（单路件）分工：单路去抖归
 *                         那件、16 路批量库归本件；与 `FB_DL_PulseWidthFilter`
 *                         分工：脉宽滤除 ≠ 电平去抖。
 * 来源标签 (Source Tag) : IEC 61131-3 标准语义的道莅防御性实现（TON 双阈值
 *                         去抖为标准定时器语义组合）
 * 码表     (Codes)      : 本件不占用任何全局数字码位。出口为 BOOL 数组 +
 *                         ENUM 信息码；数字码位待主控收口阶段统一派号。
 * 红线自检 (Redline)    : R1 ✓ 零 GVL/VAR_EXTERNAL ｜ R2 ✓ 零 %I/%Q/%M ｜ R3 ✓ 纯 IEC 61131-3
 *                         R4 ✓ 通道钳位 + 时间域兜底 + 有效域外恒 FALSE ｜ R5 ✓ 声明逐行同行双语注释
 *                         R6 N/A（无 ENUM 状态机） ｜ R7 ✓ 32 TON 段 0 定长循环无条件刷新
 * 修订历史 (Revision)   : 2026-11-20  v1.0.0  R50 首版（批次 1 · 序号 4）
 * 验收向量 (Acceptance) : ① 通道 0：tRise=T#50MS，tFall=T#50MS，原始信号跳变
 *                         TRUE 后 30ms 输出仍 FALSE（确认窗内保持），50ms 后
 *                         abDeb[0]=TRUE；② 原始信号 20ms 毛刺（< 50ms）：输出
 *                         不翻转（毛刺被去抖）；③ nChanCnt=20 → 钳位 16，
 *                         eErrCode=eCfgClamp；nChanCnt=0 → 钳位 1，
 *                         eErrCode=eCfgClamp，通道 1~15 恒 FALSE。
 *==============================================================================*)

(*-----------------------------------------------------------------------------
 * 枚举: E_DL_DbbErr（信息码；钳位走信息级，不置 bError）
 *----------------------------------------------------------------------------*)
TYPE E_DL_DbbErr :
(
    eOk       := 0,   // 通道数在合法域 / Channel count in domain
    eCfgClamp := 1    // 信息级：通道数越界已钳位 [1,16] / Info: channel count clamped to [1,16]
);
END_TYPE

FUNCTION_BLOCK FB_DL_DebounceBank
VAR_INPUT
    abRaw    : ARRAY[0..15] OF BOOL;   // 16 路原始输入信号 [-] / Sixteen raw input signals
    aRise    : ARRAY[0..15] OF TIME;   // 16 路上升确认时间（<=T#0S 直通） [ms] / Sixteen rise confirm times
    aFall    : ARRAY[0..15] OF TIME;   // 16 路下降确认时间（<=T#0S 直通） [ms] / Sixteen fall confirm times
    nChanCnt : UDINT := 16;            // 有效通道数，域 [1,16]（越界钳位） [路] / Active channel count
END_VAR
VAR_OUTPUT
    abDeb    : ARRAY[0..15] OF BOOL;   // 16 路去抖输出（有效域外恒 FALSE） [-] / Sixteen debounced outputs
    bStable  : BOOL;                   // 全有效通道稳定指示（无通道在确认窗内） [-] / All-active-channels stable indicator
    eErrCode : E_DL_DbbErr;            // 信息码出口 / Info code outlet
    bError   : BOOL;                   // 故障标志（本件恒 FALSE，契约位） [-] / Error flag, contract pin, always FALSE
END_VAR
VAR
    _nCount  : DINT;                   // 钳位后有效通道数 [路] / Clamped active channel count
    _bClamp  : BOOL;                   // 本拍发生钳位 [-] / Clamp occurred this scan
    _bAllStb : BOOL;                   // 稳定指示内部量 [-] / Stable indicator internal
    i        : DINT;                   // 通道循环索引 / Channel loop index
    aTonRise : ARRAY[0..15] OF TON;    // 16 路上升确认定时器（段 0 定长循环无条件调用） / Sixteen rise TON instances
    aTonFall : ARRAY[0..15] OF TON;    // 16 路下降确认定时器（段 0 定长循环无条件调用） / Sixteen fall TON instances
END_VAR
VAR CONSTANT
    DL_DBB_NMAX : DINT := 16;          // 通道定长上限 [路] / Fixed channel ceiling
    DL_DBB_NMIN : DINT := 1;           // 通道数下限 [路] / Active count floor
END_VAR

(* —— 段 0：通道数钳位 + 32 TON 定长循环无条件刷新（R6/R7） —— *)
_bClamp := FALSE;                                   // 钳位量预清 / Clamp preset
_nCount := UDINT_TO_DINT(nChanCnt);                 // 通道数转 DINT（越界由下步钳位） / Convert count
IF _nCount > DL_DBB_NMAX THEN
    _nCount := DL_DBB_NMAX;                         // 上越界钳 16 / Clamp high to 16
    _bClamp := TRUE;                                // 记钳位 / Mark clamp
END_IF
IF _nCount < DL_DBB_NMIN THEN
    _nCount := DL_DBB_NMIN;                         // 下越界钳 1 / Clamp low to 1
    _bClamp := TRUE;                                // 记钳位 / Mark clamp
END_IF
FOR i := 0 TO (DL_DBB_NMAX - 1) DO
    aTonRise[i](IN := abRaw[i],  PT := aRise[i]);   // 上升确认 TON 无条件调用 / Rise TON unconditional call
    aTonFall[i](IN := NOT abRaw[i], PT := aFall[i]);   // 下降确认 TON 无条件调用 / Fall TON unconditional call
END_FOR

(* —— 段 1：双阈值去抖输出（有效通道：Rise.Q 置 / Fall.Q 复 / 窗内保持；域外恒 FALSE） —— *)
_bAllStb := TRUE;                                   // 稳定指示起步为真，逐通道合取 / Stable preset true, AND-reduce
FOR i := 0 TO (DL_DBB_NMAX - 1) DO
    IF i >= _nCount THEN
        abDeb[i] := FALSE;                          // 有效域外通道恒 FALSE（规格④） / Out-of-domain channel constant FALSE
    ELSIF aTonRise[i].Q THEN
        abDeb[i] := TRUE;                           // 上升确认到：置 TRUE（已确认通道不降低稳定指示） / Rise confirmed: TRUE
    ELSIF aTonFall[i].Q THEN
        abDeb[i] := FALSE;                          // 下降确认到：回 FALSE / Fall confirmed: FALSE
    ELSE
        _bAllStb := FALSE;                          // 双窗均未到：输出保持上拍，本通道不稳定 / Both windows pending: hold, unstable
        (* abDeb[i] 不赋值 = 保持上拍（互斥保持语义，头注释③） *)
    END_IF
END_FOR

(* —— 段 2：出口单点映射（名实双出口同源，R191） —— *)
bStable := _bAllStb;                                // 稳定指示出口 / Stable indicator outlet
IF _bClamp THEN
    eErrCode := E_DL_DbbErr.eCfgClamp;              // 信息级：钳位口径 / Info: clamped
ELSE
    eErrCode := E_DL_DbbErr.eOk;                    // 正常 / Normal
END_IF
bError := FALSE;                                    // 本件无故障级条件（头注释声明） / No fault-level condition

END_FUNCTION_BLOCK

(* ---- FB_DL_DiagTextLookup.st ---- *)
(*==============================================================================
 * 组件名称 (Component)  : FB_DL_DiagTextLookup
 * 所属子库 (Sublibrary) : DL_Base
 * 当前版本 (Version)    : 1.0.0
 * 兼容性   (Platform)   : CODESYS 3.5 / TwinCAT 3 / 汇川 InoProShop / Machine Expert
 *                         仅依赖 Standard.library（LEN / SHR / 类型转换），零厂商方言
 * 来源标签 (Source)     : self-std
 * 功能描述 (Function)   : 诊断码到 HMI 文本的纯查表：32 位诊断码低 16 位为表内下标，
 *                         高 16 位为段位（0001 / 0003 等分段路由信息，原样导出给 HMI）。
 *                         命中返回该行文本（中英双数组，按语言选择位取一）；
 *                         未命中返回空串占位行并置 bNotFound；文本超 255 字符按
 *                         R49 四步样板先置截断码再钳长写入。
 *                         每拍重算不锁存（纯查表语义，规格明示：本件无时序状态机，
 *                         故障级码同为每拍重算，规格条款优先于锁存惯例）。
 * 边界与语义披露 (Boundary disclosure) :
 *   1) 文本数组经 VAR_IN_OUT 注入（零全局耦合）：中英两数组维度一致 [0..63]、
 *      元素 STRING(512)——源行允许长于输出上限，截断防御真实可达；
 *      输出 sText / sTextOpp 固定 STRING(255)。
 *   2) 码位高段掩码路由：nIdx = 低 16 位掩码 AND 的无符号值，段位不参与寻址；
 *      段位经 uSegment 原样导出（0001 = Base 族、0003 = Device 族等），HMI 据此分组。
 *   3) 未命中（下标越出有效行数）与组态非法（表长 <= 0）输出不同的码位与标志：
 *      未命中为信息级 + bNotFound，组态非法为故障级 + bError + 输出空串。
 *   4) 本件无定时器 / 无边沿 / 无状态驻留：每拍纯重算，失能语义即组态非法语义。
 * 故障码表 (Error codes) :
 *   16#0001_03F2 [故障级] 表长组态非法（<1 或 >64），输出空串 + bNotFound + bError
 *                 反证：该场景输出空串且 bNotFound 置位，与「未命中」输出组合
 *                 完全相同，无故障级码则组态错误会被当成普通未命中静默放过。
 *   16#0001_04B6 [信息级] 码位未命中（下标越出有效行数），返回空串占位行
 *                 反证：bNotFound 已置位，但 HMI 事件流水需要码位归档未命中
 *                 频次（高频未命中 = 表维护缺失），布尔位不承载频次。
 *   16#0001_04B7 [信息级] 命中行文本超 255 字符，已按 R49 先置码后钳长
 *                 反证：截断后的文本与真实 255 长文本输出组合相同，无码则
 *                 截断事实不可观测（R49 截断码赋值行先于钳位行，本件已按序）。
 * 码位总账 (Code ledger) : 16#0001_03F2 用 ｜ 16#0001_04B6 / 04B7 用
 * 依赖     (Depends)    : 无 DL_ 内部依赖；Standard.library: LEN / SHR
 * 红线自检 (Redline)    : R1 ✓ 零全局变量与 VAR_EXTERNAL ｜ R2 ✓ 零 %I/%Q 物理地址
 *                         R3 ✓ 纯 IEC 61131-3 ｜ R4 ✓ 表长域闸 / 下标界检（LOWER/UPPER 口径）
 *                         R5 ✓ 全变量中英双语同行注释 ｜ R6 N/A（纯查表，无状态机无 CASE）
 *                         R7 N/A（无定时器 / 边沿实例）
 * 修订历史 (Revision)   :
 *   2026-11-22  v1.0.0  首版入库（R68 构建轮 · 批 1 · 目标 3）
 *============================================================================*)
FUNCTION_BLOCK FB_DL_DiagTextLookup
VAR_INPUT
    uCodeIn    : UDINT := 0;    // 输入诊断码 [码]，低 16 位 = 表内下标 / Diagnostic code in, low word = index
    nTableLen  : INT   := 64;   // 有效行数 [行]，域 1..64，越界组态非法 / Valid row count, 1..64
    bEnglish   : BOOL  := FALSE;// 语言选择位：FALSE = 中文，TRUE = 英文 / Language select, FALSE Chinese
    bEnable    : BOOL  := TRUE; // 查表使能（FALSE 输出空串安全态）/ Lookup enable, FALSE safe empty
END_VAR
VAR_IN_OUT
    azhTable : ARRAY[0..63] OF STRING(512);  // 中文文本表 [0..63 行]，注入引用 / Chinese text table, injected by reference
    aenTable : ARRAY[0..63] OF STRING(512);  // 英文文本表 [0..63 行]，注入引用 / English text table, injected by reference
END_VAR
VAR_OUTPUT
    sText      : STRING(255);   // 命中文本（按语言选择位）/ Hit text per the language select
    sTextOpp   : STRING(255);   // 另一语言文本（双语 HMI 诊断用）/ Text in the other language
    bNotFound  : BOOL;          // 未命中标志（本拍重算）/ Not found flag, recomputed every scan
    bTruncated : BOOL;          // 截断标志（本拍重算，R49 先码后钳）/ Truncated flag, code set before clamp
    uSegment   : UDINT;         // 码位高段（0001 / 0003 等分段路由）/ High segment of the code for routing
    bError     : BOOL;          // 故障标志（表长组态非法，每拍重算）/ Fault flag, config class
    uErrorId   : UDINT;         // 故障码，0 = 无故障（每拍重算）/ Error code, recomputed every scan
    bValid     : BOOL;          // 本拍查表有效命中 / A valid hit this scan
END_VAR
VAR
    nIdx      : DINT;           // 低 16 位下标 [行]，DINT 承载防 0xFFFF 越界 INT / Low-word index as DINT
    sSrcSel   : STRING(512);    // 选中语言源行快照 / Selected language source row snapshot
    sSrcOpp   : STRING(512);    // 另一语言源行快照 / Other language source row snapshot
    bHit      : BOOL;           // 本拍下标命中 / Index hit this scan
    nLenSel   : INT;            // 选中行长度 [字符]，LEN 标准返回 INT / Selected row length, LEN returns INT
    nLenOpp   : INT;            // 另一语言行长度 [字符] / Other row length
END_VAR
VAR CONSTANT
    DL_DT_IDX_MASK : UDINT := 16#0000_FFFF;  // 低 16 位下标掩码 / Low-word index mask
    DL_DT_SEG_SHFT : UDINT := 16;            // 段位右移量 [bit]（< 32，结构性安全）/ Segment shift, structurally safe
    DL_DT_ROWS_MAX : INT   := 64;            // 表容量上限 [行]，与数组维度一致 / Table capacity, matches the arrays
    DL_DT_TEXT_MAX : INT   := 255;           // 输出文本上限 [字符]，LEN 同型 INT / Output text ceiling, INT like LEN
END_VAR

(*------------------------------------------------------------------------------
 * 段 1｜每拍预清（单拍 / 信息位统一出口预置，FB51-8①）
 *      Per-scan preset of all single-scan and info outputs
 *-----------------------------------------------------------------------------*)
sText      := '';
sTextOpp   := '';
bNotFound  := FALSE;
bTruncated := FALSE;
bValid     := FALSE;
bError     := FALSE;
uErrorId   := 16#0000_0000;
uSegment   := 16#0000_0000;

(*------------------------------------------------------------------------------
 * 段 2｜组态域闸（R151）：表长 <1 或 >64 即非法，输出安全态（空串）
 *      Config gate: table length out of 1..64 is illegal, safe empty output
 *      组态非法为结构性分支（IF/ELSE 全覆盖），不用 RETURN 早退（失能路径清输出）
 *-----------------------------------------------------------------------------*)
IF (NOT bEnable) OR (nTableLen < 1) OR (nTableLen > DL_DT_ROWS_MAX) THEN
    (* 组态非法 / 失能：空串安全态 + 故障级码（失能与非法共用安全出口，码位区分） *)
    (* Illegal or disabled: safe empty output, fault code tells the two apart *)
    IF (nTableLen < 1) OR (nTableLen > DL_DT_ROWS_MAX) THEN
        uErrorId := 16#0001_03F2;   // 故障级：表长组态非法 / Fault: table length illegal
        bError   := TRUE;           // R45 配对 / Paired with the fault code
        bNotFound := TRUE;          // 非法态同样视为未命中语义 / Illegal also means not found
    END_IF
ELSE
    (*------------------------------------------------------------------------------
     * 段 3｜下标路由与段位导出（边界 B2）
     *      Index routing and segment export
     *      UDINT_TO_DINT：0xFFFF = 65535 超出 INT 正域，必须升位 DINT 承载（R55）
     *-----------------------------------------------------------------------------*)
    nIdx    := UDINT_TO_DINT(uCodeIn AND DL_DT_IDX_MASK);
    uSegment := SHR(uCodeIn, DL_DT_SEG_SHFT);
    bHit    := (nIdx >= 0) AND (nIdx < UDINT_TO_DINT(nTableLen));

    IF bHit THEN
        (*------------------------------------------------------------------------------
         * 段 4｜命中：双语言取行 + R49 四步截断样板
         *      Hit: fetch both rows, R49 four-step truncation template
         *      步 1 测长 -> 步 2 超限置码 -> 步 3 钳长（赋值即钳） -> 步 4 写出
         *      步 1 measure, step 2 code, step 3 clamp by assignment, step 4 write
         *-----------------------------------------------------------------------------*)
        IF bEnglish THEN
            sSrcSel := aenTable[DINT_TO_INT(nIdx)];
            sSrcOpp := azhTable[DINT_TO_INT(nIdx)];
        ELSE
            sSrcSel := azhTable[DINT_TO_INT(nIdx)];
            sSrcOpp := aenTable[DINT_TO_INT(nIdx)];
        END_IF

        nLenSel := LEN(sSrcSel);        // 标准 LEN 返回 INT / Standard LEN returns INT
        nLenOpp := LEN(sSrcOpp);

        IF nLenSel > DL_DT_TEXT_MAX THEN
            bTruncated := TRUE;          // 步 2 截断码先行（R49：码先于钳）/ Code before clamp
            uErrorId   := 16#0001_04B7;
        END_IF
        IF nLenOpp > DL_DT_TEXT_MAX THEN
            bTruncated := TRUE;          // 另一语言超限同置标志 / Other language truncation too
            IF uErrorId = 16#0000_0000 THEN
                uErrorId := 16#0001_04B7;
            END_IF
        END_IF

        sText    := sSrcSel;             // 步 3+4：赋值即按 255 钳长写出 / Clamp by assignment
        sTextOpp := sSrcOpp;
        bValid   := TRUE;
    ELSE
        (*------------------------------------------------------------------------------
         * 段 5｜未命中：空串占位行 + 信息级码（每拍重算，不锁存）
         *      Miss: empty placeholder row plus info code, recomputed per scan
         *-----------------------------------------------------------------------------*)
        sText     := '';
        sTextOpp  := '';
        bNotFound := TRUE;
        uErrorId  := 16#0001_04B6;
    END_IF
END_IF
END_FUNCTION_BLOCK

(* ---- FB_DL_DualEdgeTrig.st ---- *)
(*==============================================================================
 * 组件名称 (Component)  : FB_DL_DualEdgeTrig
 * 所属子库 (Sublibrary) : DL_Base
 * 当前版本 (Version)    : 1.0.1
 * 兼容性   (Platform)   : CODESYS 3.5 / TwinCAT 3 / 汇川 InoProShop / Machine Expert
 *                         仅依赖 Standard.library（R_TRIG），零厂商方言
 * 功能描述 (Function)   : 双边沿检测器。同一实例一次给出上升沿 / 下降沿 / 任意跳变
 *                         三种单扫描周期脉冲与当前电平，并累计上升/下降次数。
 *                         替代"一处用 R_TRIG、另一处用 NOT 取下降沿"的散乱写法，
 *                         统一多工位取沿的语义。计数器达上限后饱和停增并告警（不回绕）。
 * 开源溯源 (Origin)     : 原创实现。语义参照 IEC 61131-3 标准 R_TRIG 定义与
 *                         PLCopen Coding Guidelines 的单一事件源原则。
 * 依赖     (Depends)    : 无 DL_ 内部依赖；Standard.library: R_TRIG
 * 红线自检 (Redline)    : R1 ✓ 零全局变量表与外部变量引用 ｜ R2 ✓ 零物理 IO 地址直写
 *                         R3 ✓ 纯 IEC 61131-3 ｜ R4 ✓ 计数饱和+首扫抑制
 *                         R5 ✓ 全变量中英双语同行注释 ｜ R6 N/A（无边沿无关状态机，见下）
 *                         R7 ✓ 三实例主体最前部无条件刷新
 * 说明     (Note)       : R6 标注 N/A —— 本组件不存在顺序状态机，仅为边沿锁存与计数，
 *                         无 CASE 可写；非法状态不可能出现（唯一状态即"运行"），
 *                         故以本节说明替代 ELSE 兜底，符合 R6"无状态机则标注 N/A"口径。
 * 修订历史 (Revision)   :
 *   2026-11-14  v1.0.0  首版入库（Phase 1 冷启动 · Level 0 批次）
 *   2026-11-14  v1.0.1  修复事件校正极性反接缺陷：上升/下降两路的事件
 *                       与"上一周期电平"的与项被写反，导致真实跳变周期被自身屏蔽、
 *                       两个事件输出恒为 FALSE（计数永不增长）。改为上升沿与
 *                       "上周期为低"相与、下降沿与"上周期为高"相与，与
 *                       bLastLevel 的更新时机（事件判定之后）保持一致。
 *============================================================================*)
FUNCTION_BLOCK FB_DL_DualEdgeTrig
VAR_INPUT
    bSignal    : BOOL;            // 待检测信号，建议已消抖 / Signal to detect, pre-debounced recommended
    bEnable    : BOOL := TRUE;    // 使能标志，FALSE 时所有事件强制 FALSE / Enable flag, FALSE forces all events FALSE
    bReset     : BOOL;            // 复位信号，上升沿清零计数器并抑制当周期事件 / Reset, rising edge clears counters and suppresses events
END_VAR
VAR_OUTPUT
    bLevel     : BOOL;            // 当前电平，始终直通 / Current level, always pass-through
    bRising    : BOOL;            // 上升沿，单扫描周期脉冲 / Rising edge, one-scan pulse
    bFalling   : BOOL;            // 下降沿，单扫描周期脉冲 / Falling edge, one-scan pulse
    bChanged   : BOOL;            // 任意跳变 = 上升 OR 下降 / Any transition = rising OR falling
    uRiseCount : UDINT;           // 累计上升沿次数 / Accumulated rising edge count
    uFallCount : UDINT;           // 累计下降沿次数 / Accumulated falling edge count
    uErrorId   : UDINT;           // 故障码，仅计数器饱和告警 / Error code, counter saturation warning only
END_VAR
VAR
    fbTrigRise  : R_TRIG;         // 上升沿检测实例 / Rising edge detector instance
    fbTrigFall  : R_TRIG;         // 下降沿检测实例，输入取反信号 / Falling edge detector instance on inverted signal
    fbTrigReset : R_TRIG;         // 复位信号上升沿检测实例 / Reset rising edge detector instance
    bLastLevel  : BOOL;           // 上一周期电平，用于事件校正 / Previous level, used for event qualification
    bFirstScan  : BOOL := TRUE;   // 上电首扫标志，TRUE 期间抑制全部事件 / First-scan flag, suppresses all events while TRUE
END_VAR
VAR CONSTANT
    DL_EDGE_COUNT_MAX : UDINT := 16#FFFF_FFFE;  // 计数饱和上限，达上限停增不回绕 / Counter saturation limit, no wrap-around
END_VAR

(*------------------------------------------------------------------------------
 * 段 1｜无条件刷新区（红线 R7）：三个 R_TRIG 实例严禁进入任何 IF / CASE 分支
 *      Unconditional refresh zone (red line R7): no instance call inside IF / CASE
 *      下降沿走"取反信号"的对称路径，避免手写 IF NOT 分支时漏掉首扫抑制
 *-----------------------------------------------------------------------------*)
fbTrigRise(CLK := bSignal);
fbTrigFall(CLK := NOT bSignal);
fbTrigReset(CLK := bReset);

IF bFirstScan THEN
    (*--------------------------------------------------------------------------
     * 段 2｜上电首扫（边界 B2）：同步电平与历史电平，三类事件全部清零
     *      R_TRIG 首扫本身可能因 CLK 为 TRUE 而输出 Q，故必须显式抑制一周期
     *      First scan: synchronize levels and clear all events explicitly
     *-------------------------------------------------------------------------*)
    bLevel     := bSignal;
    bLastLevel := bSignal;
    bRising    := FALSE;
    bFalling   := FALSE;
    bChanged   := FALSE;
    bFirstScan := FALSE;
ELSE

    (* 段 3｜电平直通：使能关闭时电平仍必须真实反映输入（边界 B6） *)
    (* Level pass-through: level must stay truthful even when disabled (boundary B6) *)
    bLevel := bSignal;

    IF fbTrigReset.Q THEN
        (*----------------------------------------------------------------------
         * 段 4｜复位语义（边界 B5）：清计数、抑制当周期事件、同步历史电平
         *      Reset: clear counters, suppress current-scan events, resync last level
         *---------------------------------------------------------------------*)
        uRiseCount := 16#0000_0000;
        uFallCount := 16#0000_0000;
        uErrorId   := 16#0000_0000;
        bRising    := FALSE;
        bFalling   := FALSE;
    ELSE
        IF bEnable THEN
            (*------------------------------------------------------------------
             * 段 5｜事件判定（边界 B1/B3）：R_TRIG 的 Q 再与上一周期电平做校正
             *      校正的目的：实例被跨任务共享或重复调用时 bLastLevel 尚未建立，
             *      单靠 Q 会把"初始电平"误当成一次跳变
             *      Event qualification: Q is AND-ed with the previous level
             *      极性口径（v1.0.1 修正）：真实上升沿那一周期 bLastLevel 必为 FALSE，
             *      故上升沿与 NOT bLastLevel 相与；下降沿取反信号做 CLK，
             *      跳变周期 bLastLevel 必为 TRUE，故下降沿与 bLastLevel 相与。
             *      上一版两路极性接反，跳变周期被自身屏蔽，事件恒不成立。
             *      Polarity: a rise implies the previous level was low, and the
             *      falling path clocks on the inverted signal, so its previous
             *      level is high. v1.0.1 corrects the two qualifiers that were swapped.
             *-----------------------------------------------------------------*)
            bRising  := fbTrigRise.Q AND NOT bLastLevel;
            bFalling := fbTrigFall.Q AND bLastLevel;
        ELSE
            (* 使能关闭：事件全部清零，但历史电平在本段末尾继续跟踪（边界 B6） *)
            (* Disabled: clear all events, yet last level keeps tracking at the end of this block *)
            bRising  := FALSE;
            bFalling := FALSE;
        END_IF

        IF bRising THEN
            (*------------------------------------------------------------------
             * 段 6｜上升计数：饱和停增，禁止回绕归零（边界 B4）
             *      Rising count: saturate at limit, wrap-around is forbidden
             *-----------------------------------------------------------------*)
            IF uRiseCount < DL_EDGE_COUNT_MAX THEN
                uRiseCount := uRiseCount + 1;
            ELSE
                uErrorId := 16#0001_0007;
            END_IF
        END_IF

        IF bFalling THEN
            (*------------------------------------------------------------------
             * 段 7｜下降计数：与上升计数同一饱和策略，保证两路对称
             *      Falling count: identical saturation policy for symmetry
             *-----------------------------------------------------------------*)
            IF uFallCount < DL_EDGE_COUNT_MAX THEN
                uFallCount := uFallCount + 1;
            ELSE
                uErrorId := 16#0001_0007;
            END_IF
        END_IF
    END_IF

    (* 段 8｜跳变合成：bChanged 由两路事件或运算得到，天然互斥（边界 B3） *)
    (* Transition composition: bChanged is the OR of both events, mutually exclusive by nature *)
    bChanged := bRising OR bFalling;

    (* 段 9｜历史电平更新：必须放在事件判定之后，且禁用时也执行（边界 B6） *)
    (* Last level update: must follow event evaluation and also runs while disabled *)
    bLastLevel := bSignal;
END_IF
END_FUNCTION_BLOCK

(* ---- FB_DL_DualWindowBandCmp.st ---- *)
// FB_DL_DualWindowBandCmp v1.0.0
// 开源溯源：brOscatLib / URL https://github.com/iec-oscat-mirror / 许可证 MIT / 借鉴 WINDOW2 双窗三态语义，clean-room 重写
(*
  道莅工业代码库 | DL_Base | FB_DL_DualWindowBandCmp
  版本: 1.0.0 | 日期: 2026-11-23 | 轮次: R75
  功能: 双独立窗口三态比较器（下窗/带内/上窗），窗口 A/B 各自独立判定，
        并输出双窗一致性（同带）判据
  邻件关系: 与 FC_DL_ToleranceWindow（单容差窗布尔判定）相邻 —— 差异点：
            容差窗为单窗带内/带外两态布尔，本件为双窗各三态枚举 + 同带
            一致性输出，语义扩展非同义替换
*)
TYPE E_DL_WindowBand3 :
(
    eBelow  := 0,    // 低于窗下限 / Below window low limit
    eInBand := 10,   // 带内 / Within band
    eAbove  := 20    // 高于窗上限 / Above window high limit
);
END_TYPE

FUNCTION_BLOCK FB_DL_DualWindowBandCmp
VAR_INPUT
    fValA    : REAL := 0.0;                      // 窗 A 判定值 [工程单位] / Window A value
    fLowA    : REAL := 0.0;                      // 窗 A 下限 [工程单位] / Window A low limit
    fHighA   : REAL := 100.0;                    // 窗 A 上限 [工程单位] / Window A high limit
    fValB    : REAL := 0.0;                      // 窗 B 判定值 [工程单位] / Window B value
    fLowB    : REAL := 0.0;                      // 窗 B 下限 [工程单位] / Window B low limit
    fHighB   : REAL := 100.0;                    // 窗 B 上限 [工程单位] / Window B high limit
    fEps     : REAL := 1.0E-6;                   // 浮点判等容差 [工程单位] / Float equality tolerance
END_VAR
VAR_OUTPUT
    eBandA     : E_DL_WindowBand3;               // 窗 A 三态判定 / Window A three-state band
    eBandB     : E_DL_WindowBand3;               // 窗 B 三态判定 / Window B three-state band
    bBothIn    : BOOL;                           // 双窗同时带内 [-] / Both windows in band
    bSameBand  : BOOL;                           // 双窗同带（枚举相等）[-] / Same band on both windows
    bValid     : BOOL;                           // 组态有效回执 [-] / Configuration validity receipt
    bError     : BOOL;                           // 故障标志（组态非法）/ Fault flag (invalid configuration)
    uErrorId   : UDINT;                          // 事件码，0 = 无事件；16#0002_1C01 = 窗限组态非法 / Event code
END_VAR

// —— 段 0：全路径缺省 —— //
eBandA := E_DL_WindowBand3.eInBand;              // 三态缺省带内（安全中性值）/ Default neutral in-band
eBandB := E_DL_WindowBand3.eInBand;              // 窗 B 缺省 / Window B default
bBothIn := FALSE;                                // 一致性预清 / Agreement preset
bSameBand := FALSE;                              // 同带预清 / Same-band preset
bValid := FALSE;                                 // 有效回执预清 / Validity preset
bError := FALSE;                                 // 故障预清（组态非法路径置位）/ Fault preset
uErrorId := 16#0000;                             // 事件码预清 / Event code preset

// —— 段 1：组态闸（窗限单调 + 非有限 + 容差非负） —— //
IF (fLowA > fHighA + fEps) OR (fLowB > fHighB + fEps) THEN   // 窗限倒置（容差判等）/ Window limits inverted
    bError := TRUE;                              // 故障级：组态非法 / Fault level: invalid config
    uErrorId := 16#0002_1C01;                    // 故障码（1Cxx 步进）/ Fault code
    RETURN;                                      // 非法组态不判定 / No judgment on invalid config
END_IF
IF (fValA <> fValA) OR (fValB <> fValB) OR (fLowA <> fLowA) OR (fHighA <> fHighA)
   OR (fLowB <> fLowB) OR (fHighB <> fHighB) THEN
    bError := TRUE;                              // 任一输入 NaN / Any input NaN
    uErrorId := 16#0002_1C01;                    // 同组态故障码 / Same fault code family
    RETURN;
END_IF
bValid := TRUE;                                  // 组态与输入均有效 / Config and inputs valid

// —— 段 2：窗 A 三态判定（带界按闭区间，容差判等） —— //
IF fValA < fLowA - fEps THEN                     // 低于下限（容差外）/ Below low with tolerance
    eBandA := E_DL_WindowBand3.eBelow;
ELSIF fValA > fHighA + fEps THEN                 // 高于上限（容差外）/ Above high with tolerance
    eBandA := E_DL_WindowBand3.eAbove;
ELSE                                             // 带内（含边界容差带）/ Within band incl. boundary
    eBandA := E_DL_WindowBand3.eInBand;
END_IF

// —— 段 3：窗 B 三态判定（同口径） —— //
IF fValB < fLowB - fEps THEN                     // 窗 B 低于下限 / Window B below low
    eBandB := E_DL_WindowBand3.eBelow;
ELSIF fValB > fHighB + fEps THEN                 // 窗 B 高于上限 / Window B above high
    eBandB := E_DL_WindowBand3.eAbove;
ELSE                                             // 窗 B 带内 / Window B in band
    eBandB := E_DL_WindowBand3.eInBand;
END_IF

// —— 段 4：一致性输出（双窗同带 + 双带内） —— //
bBothIn := (eBandA = E_DL_WindowBand3.eInBand) AND (eBandB = E_DL_WindowBand3.eInBand);   // 双带内 / Both in band
bSameBand := (eBandA = eBandB);                  // 枚举相等判同带（浮点禁等令不适用于枚举）/ Same band by enum equality
END_FUNCTION_BLOCK

(* ---- FB_DL_DutyCycleMeasure.st ---- *)
(*
  ==================================================================
  组件名 Component  : FB_DL_DutyCycleMeasure
  分类   Category   : DL_Base
  版本   Version    : 1.0.0
  功能   Purpose    : 占空比/周期双沿测量：上升沿→上升沿累计测周期，高电平
                      期间累计测高宽度，周期闭合拍一次性算占空比并钳位 0~100。
                      首周期未闭合不出数（bValid=FALSE）；闭合周期累计值 ≤ 0
                      视为无效测量，bValid=FALSE 且保持上次输出值（不静默清零）。
                      周期闭合判据用「累计值 > 0」整数级事实，禁浮点判等。
  来源   Source     : t2-1-lgf-measurement（测量族：双沿计时口径为公开教科书
                      算法，实现零源码复制）
  互引   Cross-ref  : FB_DL_FrequencyGenerator（对偶件：本件测周期，彼件产生
                      频率信号，可组成环路自检）；FC_DL_PeriodJitterCalc（下游
                      可把本件 fPeriodMs 序列喂给它算抖动）
  平台   Platform   : 纯 IEC 61131-3（R_TRIG/F_TRIG/LREAL 四则），三平台通用
  依赖   Depends    : 仅 Standard.library（R_TRIG/F_TRIG 属标准件）
  设计偏差 Deviation: 时间基准按本库「时间注入」纪律（R 平台时刻函数拒绝方案，
                      参见 FB_DL_CycleTimeMeasure 头注）：新增输入 fCallCycleMs
                      由调用方按扫描增量注入，本件不读任何平台时刻函数。
  红线   Redline    : R1 零全局/VAR_EXTERNAL/R2 零 %I/%Q/R3 纯 IEC 标准
                      R4 除法前分母 > 0 显式闸 + 输出 0~100 钳位 + 输入有限闸
                      R5 全变量双语同行注释/R6 纯时序累计无状态机（CASE 不适用）
                      R7 R_TRIG/F_TRIG 段 0 无条件刷新/R8 钳位与容差常量化
  契约   Contract   : bEnable=FALSE 语义（FB33-4 写死）：冻结全部输出保持上次
                      值、bValid=FALSE，累计器清零（失能相串清账，R 失能清账
                      条款）；重新使能从下一上升沿重新起测（首周期语义重置）。
                      fCallCycleMs ≤ 0 或非有限：本拍拒绝累计、bValid=FALSE
                      （推进判据与计时不同源防线：计时基准本身必须有效）。
  错误码 Codes      : 16#0001_0011【信息级】fCallCycleMs 非法（≤0 或非有限），
                      本拍拒绝计时
  验收   Acceptance : V1 50% 占空恒定方波 → fDutyPct≈50 ｜ V2 使能前首周期 →
                      bValid=FALSE ｜ V3 周期累计≤0 → bValid=FALSE 且保持上次
                      ｜ V4 失能 → 冻结 + 累计清零 ｜ V5 计时基准非法 → 拒绝
  变更   Revision   : 2026-11-22  v1.0.0  R66 首版（编码阶段批 1 序 2）
  ==================================================================
*)
FUNCTION_BLOCK FB_DL_DutyCycleMeasure
VAR_INPUT
    bSignal     : BOOL;               // 被测方波信号电平 [-] / the measured square wave level
    bEnable     : BOOL := FALSE;      // 使能，FALSE 冻结输出并清累计（头注契约）[-] / the enable, false freezes outputs and clears accumulators
    fCallCycleMs: LREAL := 0.0;       // 调用方注入的扫描周期增量 [ms] / caller injected scan delta [ms]
END_VAR
VAR_OUTPUT
    fPeriodMs   : LREAL := 0.0;       // 最近一次闭合周期 [ms]（无效拍保持上次值）/ the last closed period [ms], held when invalid
    fDutyPct    : LREAL := 0.0;       // 最近一次闭合占空比，钳位 0~100 [%]（无效拍保持）/ the last closed duty, clamped 0 to 100 [%], held when invalid
    bValid      : BOOL := FALSE;      // 本拍输出有效标志（首周期未闭合=FALSE）[-] / the output validity, false until the first period closes
    uErrorId    : UDINT := 16#0000_0000; // 错误码，0=正常，16#0001_0011=计时基准非法 [码] / the error code [code]
END_VAR
VAR
    rtSig       : R_TRIG;             // 信号上升沿实例，段 0 无条件刷新 / the rising edge instance refreshed unconditionally
    ftSig       : F_TRIG;             // 信号下降沿实例，段 0 无条件刷新 / the falling edge instance refreshed unconditionally
    _bHasEdge   : BOOL := FALSE;      // 首个上升沿是否已捕获（FALSE=首周期未闭合）[-] / the first rising edge captured flag
    _fCycAccMs  : LREAL := 0.0;       // 当前周期累计时长 [ms] / the current period accumulator [ms]
    _fHiAccMs   : LREAL := 0.0;       // 当前周期高电平累计时长 [ms] / the current high level accumulator [ms]
    _bTimeOk    : BOOL := FALSE;      // 本拍计时基准有效性 [-] / the per scan time base validity
END_VAR
VAR CONSTANT
    DCM_DUTY_MIN : LREAL := 0.0;      // 占空比输出下限 [%] / duty output lower clamp [%]
    DCM_DUTY_MAX : LREAL := 100.0;    // 占空比输出上限 [%] / duty output upper clamp [%]
    DCM_ERR_TIME : UDINT := 16#0001_0011; // 计时基准非法（信息级）/ invalid time base, info level
    DCM_ERR_NONE : UDINT := 16#0000_0000; // 无错误 [码] / no error [code]
END_VAR

(*------------------------------------------------------------------------------
 * 段 0｜沿检测无条件刷新区（红线 R7）：严禁移入 IF / CASE
 *      Edge instances refresh unconditionally, never inside a condition
 *-----------------------------------------------------------------------------*)
rtSig(CLK := bSignal);  // 上升沿 / the rising edge
ftSig(CLK := bSignal);  // 下降沿 / the falling edge

(*------------------------------------------------------------------------------
 * 段 1｜错误码本拍预置（当前周期事实，非锁存）
 *      The error code is a per scan fact, preset each cycle
 *-----------------------------------------------------------------------------*)
uErrorId := DCM_ERR_NONE;  // 预置无错误 / preset no error

(*------------------------------------------------------------------------------
 * 段 2｜失能相串清账：冻结输出 + bValid 撤销 + 累计器清零（R 失能清账）
 *      Disable phase clears the books: freeze outputs, revoke validity, wipe accumulators
 *-----------------------------------------------------------------------------*)
IF NOT bEnable THEN
    bValid     := FALSE;     // 失能不出数 / no output while disabled
    _bHasEdge  := FALSE;     // 首周期语义复位，重新使能从下一上升沿起测 / re-arm from the next rising edge after re-enable
    _fCycAccMs := 0.0;       // 周期累计清零 / clear the period accumulator
    _fHiAccMs  := 0.0;       // 高电平累计清零 / clear the high level accumulator
    RETURN;                  // 冻结保持 fPeriodMs / fDutyPct 上次值 / outputs hold their last values
END_IF

(*------------------------------------------------------------------------------
 * 段 3｜计时基准闸（推进判据与超时计时不得同源的计时侧防线）：
 *      ≤ 0 或非有限即拒绝本拍计时，bValid 撤销，输出保持上次值
 *      Reject the whole scan when the time base is illegal or non finite
 *-----------------------------------------------------------------------------*)
_bTimeOk := (fCallCycleMs > 0.0) AND (fCallCycleMs = fCallCycleMs);  // 自反判 NaN，> 0 排除零与负 / reflexive NaN test and positive gate
IF NOT _bTimeOk THEN
    bValid   := FALSE;          // 撤销有效性，输出保持 / revoke validity, outputs hold
    uErrorId := DCM_ERR_TIME;   // 信息级码（不置故障锁存）/ info level code, no fault latch
    _fCycAccMs := 0.0;          // 丢弃脏累计，避免混入错误时间基准的样本 / drop the dirty accumulation
    _fHiAccMs  := 0.0;          // 同上 / the same
    RETURN;
END_IF

(*------------------------------------------------------------------------------
 * 段 4｜正常计时累计：周期全程累计 + 高电平条件累计
 *      Normal accumulation: period accumulates all scan, high only when level
 *-----------------------------------------------------------------------------*)
_fCycAccMs := _fCycAccMs + fCallCycleMs;  // 周期累计 [ms] / accumulate the period [ms]
IF bSignal THEN
    _fHiAccMs := _fHiAccMs + fCallCycleMs;  // 高电平宽度累计 [ms] / accumulate the high width [ms]
END_IF

(*------------------------------------------------------------------------------
 * 段 5｜上升沿闭合周期：非首沿才出数；闭合判据为累计值 > 0，禁浮点判等
 *      A rising edge closes the period, only when it is not the first edge
 *-----------------------------------------------------------------------------*)
IF rtSig.Q THEN
    IF _bHasEdge THEN
        IF _fCycAccMs > 0.0 THEN        // 闭合判据：整数级事实「累计为正」/ close test is the positive accumulator fact
            fPeriodMs := _fCycAccMs;    // 发布闭合周期 [ms] / publish the closed period [ms]
            fDutyPct  := (_fHiAccMs / _fCycAccMs) * DCM_DUTY_MAX;  // 分母已闸 > 0 / the denominator is gated above zero
            IF fDutyPct < DCM_DUTY_MIN THEN
                fDutyPct := DCM_DUTY_MIN;   // 显式下限钳位 / explicit lower clamp
            END_IF
            IF fDutyPct > DCM_DUTY_MAX THEN
                fDutyPct := DCM_DUTY_MAX;   // 显式上限钳位 / explicit upper clamp
            END_IF
            bValid := TRUE;             // 周期闭合，输出生效 / the period closed, the outputs are live
        ELSE
            bValid := FALSE;            // 分母周期 ≤ 0：不出数且保持上次输出（头注契约）/ keep last outputs when the period is not positive
        END_IF
    END_IF
    _bHasEdge  := TRUE;   // 首沿已捕获 / the first edge is captured
    _fCycAccMs := 0.0;    // 新周期累计从零起 / the new period accumulates from zero
    _fHiAccMs  := 0.0;    // 高电平累计同步清零 / the high accumulator resets with it
END_IF
END_FUNCTION_BLOCK
